Universal Robots URScript: T013_qwen2.5-coder_32b_baseline_rep1_retry3.urscript

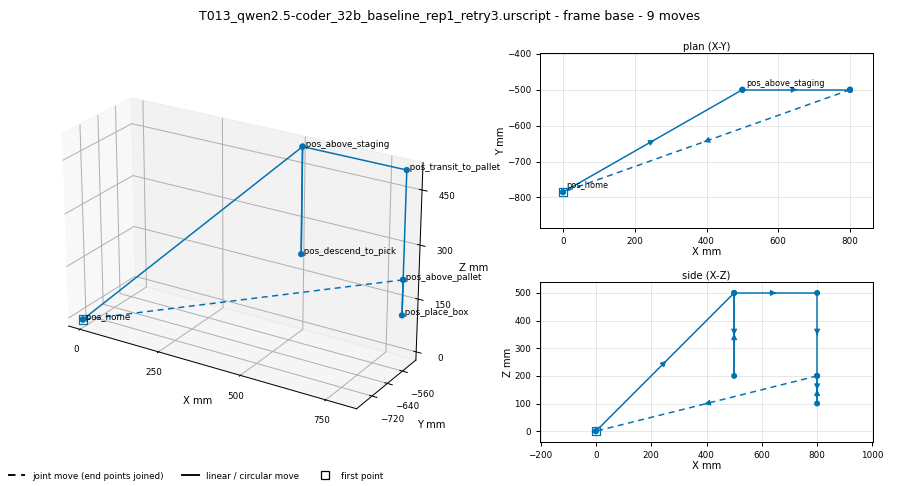
[picture p0: tool path of T013_qwen2.5-coder_32b_baseline_rep1_retry3.urscript in frame base, 9 of 9 moves have a stored position in this frame; points joined in program order, loops and branches not executed]
def collaborative_palletizing():
    # Define positions
    pos_home = p[0.0, -0.785398, 0.0, -2.356194, -1.570796, 0.0]
    pos_above_staging = p[0.5, -0.5, 0.5, 3.14, 0, 0]
    pos_descend_to_pick = p[0.5, -0.5, 0.2, 3.14, 0, 0]
    pos_lift = p[0.5, -0.5, 0.5, 3.14, 0, 0]
    pos_transit_to_pallet = p[0.8, -0.5, 0.5, 3.14, 0, 0]
    pos_above_pallet = p[0.8, -0.5, 0.2, 3.14, 0, 0]
    pos_place_box = p[0.8, -0.5, 0.1, 3.14, 0, 0]
    pos_return_above_pallet = p[0.8, -0.5, 0.2, 3.14, 0, 0]

    # Set payload
    set_payload(0.8)

    # Move to home position
    movej(pos_home, a=1.4, v=1.05, r=0)

    # Approach staging area
    movel(pos_above_staging, a=1.2, v=0.9, r=0)

    # Descend to pick box
    movel(pos_descend_to_pick, a=1.2, v=0.4, r=0)

    # Activate suction cup (simulated)
    textmsg("Activate Suction Cup")

    # Lift the box
    movel(pos_lift, a=1.2, v=0.7, r=0)

    # Transit to pallet area
    movel(pos_transit_to_pallet, a=1.3, v=0.9, r=0)

    # Approach pallet
    movel(pos_above_pallet, a=1.2, v=0.8, r=0)

    # Descend to place box
    movel(pos_place_box, a=1.2, v=0.4, r=0)

    # Deactivate suction cup (simulated)
    textmsg("Deactivate Suction Cup")

    # Lift from pallet
    movel(pos_return_above_pallet, a=1.2, v=0.7, r=0)

    # Return to home position
    movej(pos_home, a=1.4, v=1.05, r=0)
end

# Start the task
collaborative_palletizing()
